Fanuc KAREL source: KO00007.KL

PROGRAM KO00007
%NOLOCKGROUP
VAR
  P1: POSITION
  P2: POSITION
  P3: POSITION
  P4: POSITION
  OUT: XYZWPREXT
BEGIN
  OUT = FRAME(P1, P2, P3, P4)
END KO00007
